(* IEC 61131-3 sources: sigmatek-logger-api/IXON_API/Class/_TCPIPClient (part 2) *)

END_FUNCTION

FUNCTION _TCPIPClient::SendTCP
	VAR_INPUT
		pConnection 	: ^_CONNECTION;
		pData 	: ^CHAR;
		udSize 	: UDINT;
		udTimeout 	: UDINT;
	END_VAR
	VAR_OUTPUT
		dRetcode 	: DINT;
	END_VAR

  dRetcode := OS_TCP_USER_SEND(pConnection^.dSocket,
                               pData,
                               udSize,
                               0, //### flags ... not used
                               udTimeout
                               );

  if (dRetcode = udSize$DINT) then
    pConnection^.udTimeStamp := ops.tAbsolute;
  else
    udSendError += 1;
    pConnection^.FSM_TCP := _STATE_SHUTDOWN;
  end_if;

END_FUNCTION

FUNCTION _TCPIPClient::SetSocketOptions
	VAR_INPUT
		dHandle 	: DINT;
	END_VAR
	VAR_OUTPUT
		Retcode 	: DINT;
	END_VAR
VAR
	OptionValue       : DINT;
  pConn             : ^_CONNECTION;
  dRet              : DINT;
  KeepAliveLasalOS  : _KeepAliveParaLasalOS;
END_VAR

  Retcode := TCP_CLT_NO_ERROR;

  if (CheckHandleValid(dHandle) = true) then

    pConn := dHandle$^_CONNECTION;

    AP_SemaWait(AP_SemaSockOpt);

    // -----------------------------------------------------------
    // - SOCKET OPTION NAGLE
    // -----------------------------------------------------------
    if (pConn^.ConnSockOpt.Nagle = true) then
      OptionValue := 1;
    else
      OptionValue := 0;
    end_if;
    dRet := OS_TCP_USER_SETSOCKOPT(pConn^.dSocket, SOL_SOCKET, SO_NAGLE, (#OptionValue)$^CHAR, sizeof(DINT));
    if (dRet < 0) then
      Retcode := dRet;
      ConnErrCallback(pConn, TCP_CLT_ERR_GROUP_OS, dRet);
    end_if;

    // -----------------------------------------------------------
    // - SOCKET OPTION KEEP ALIVE
    // -----------------------------------------------------------
    if (bdStatus.SalamanderOS = false) then
      // --------------------------------------------------------
      // - LASAL OS
      // --------------------------------------------------------
      if (pConn^.ConnSockOpt.KeepAlive = true) then
        KeepAliveLasalOS.interval := to_UINT(pConn^.KeepAlivePara.keepIDLE);
        KeepAliveLasalOS.retry    := to_UINT(pConn^.KeepAlivePara.keepINTVL);
        KeepAliveLasalOS.timeout  := to_UINT(pConn^.KeepAlivePara.keepCNT * pConn^.KeepAlivePara.keepINTVL);
      else
        KeepAliveLasalOS.interval := 0;
        KeepAliveLasalOS.retry    := 0;
        KeepAliveLasalOS.timeout  := 0;
      end_if;
      dRet := OS_TCP_USER_SETSOCKOPT(pConn^.dSocket, SOL_SOCKET, 8, (#KeepAliveLasalOS)$^CHAR, sizeof(_KeepAliveParaLasalOS));
      if (dRet < 0) then
        Retcode := dRet;
        ConnErrCallback(pConn, TCP_CLT_ERR_GROUP_OS, dRet);
      end_if;
    else
      // --------------------------------------------------------
      // - SALAMANDER OS
      // --------------------------------------------------------
      if (pConn^.ConnSockOpt.KeepAlive = true) then
        OptionValue := 1;
      else
        OptionValue := 0;
      end_if;
      dRet := OS_TCP_USER_SETSOCKOPT(pConn^.dSocket, SOL_SOCKET, 8, (#OptionValue)$^CHAR, sizeof(DINT));
      if (dRet < 0) then
        Retcode := dRet;
        ConnErrCallback(pConn, TCP_CLT_ERR_GROUP_OS, dRet);
      end_if;

//      if (pConn^.ConnSockOpt.KeepAlive = true) then
//        OptionValue := KeepAlivePara.keepCNT;
//        dRet := OS_TCP_USER_SETSOCKOPT(pConn^.dSocket, SOL_TCP, TCP_KEEPCNT, (#OptionValue)$^CHAR, sizeof(DINT));
//        if (dRet < 0) then
//          Retcode := dRet;
//          ConnErrCallback(pConn, TCP_CLT_ERR_GROUP_OS, dRet);
//        end_if;
//        OptionValue := KeepAlivePara.keepIDLE;
//        dRet := OS_TCP_USER_SETSOCKOPT(pConn^.dSocket, SOL_TCP, TCP_KEEPIDLE, (#OptionValue)$^CHAR, sizeof(DINT));
//        if (dRet < 0) then
//          Retcode := dRet;
//          ConnErrCallback(pConn, TCP_CLT_ERR_GROUP_OS, dRet);
//        end_if;
//        OptionValue := KeepAlivePara.keepINTVL;
//        dRet := OS_TCP_USER_SETSOCKOPT(pConn^.dSocket, SOL_TCP, TCP_KEEPINTVL, (#OptionValue)$^CHAR, sizeof(DINT));
//        if (dRet < 0) then
//          Retcode := dRet;
//          ConnErrCallback(pConn, TCP_CLT_ERR_GROUP_OS, dRet);
//        end_if;
//      end_if;
    end_if;

    // -----------------------------------------------------------
    // - SOCKET OPTION DELAYED ACK
    // -----------------------------------------------------------
    if (pConn^.ConnSockOpt.DelayedAck = true) then
      OptionValue := 1;
    else
      OptionValue := 0;
    end_if;
    dRet := OS_TCP_USER_SETSOCKOPT(pConn^.dSocket, SOL_SOCKET, SO_DELAYED_ACK, (#OptionValue)$^CHAR, sizeof(DINT));
    if (dRet < 0) then
      Retcode := dRet;
      ConnErrCallback(pConn, TCP_CLT_ERR_GROUP_OS, dRet);
    end_if;

    pConn^.bdSettings.SockOptChanged := false;

    AP_SemaSignal(AP_SemaSockOpt);

  else
    Retcode := TCP_CLT_INVALID_HANDLE;
  end_if;

END_FUNCTION

FUNCTION _TCPIPClient::Read_LSLOBJ_CRC32
	VAR_INPUT
		pCRC32 	: ^CHAR;
	END_VAR
	VAR_OUTPUT
		Retcode 	: DINT;
	END_VAR
VAR
	udStrLen    : UDINT;
  udCRC32     : UDINT;
  szObjName   : ARRAY [0..255] OF CHAR;
END_VAR

  Retcode := TCP_CLT_NO_ERROR;

  if (pCRC32 <> NIL) then
    pCRC32^ := 0x00;
    udStrLen := _GetObjName(this, #szObjName[0]);
    if (udStrLen > 0) then
      udCRC32 := CheckSum.CRC32(#szObjName[0], udStrLen, 0);
      SigCLib.IToA(udCRC32$DINT, pCRC32, 0x10);
    else
      Retcode := TCP_CLT_ERR_GET_LSLOBJ_NAME;
    end_if;
  else
    Retcode := TCP_CLT_ERR_INVALID_POINTER;
  end_if;

END_FUNCTION

FUNCTION _TCPIPClient::Read_AP_TaskPeriod
	VAR_OUTPUT
		Retcode 	: DINT;
	END_VAR
VAR
	dRet          : DINT;
  LSLOBJ_INFO   : LSLOBJ_INFO;
END_VAR

  Retcode := TCP_CLT_NO_ERROR;

  dRet := _TaskObjectControl.GetObjectInfo(this, OBJ_CT, #LSLOBJ_INFO);
  case dRet of
    (*=============================================================================*)
    0: // - GET OBJECT INFO OK
    (*=============================================================================*)
      if (bdStatus.SalamanderOS = true) then
        // --------------------------------------------------------
        // - SALAMANDER OS
        // --------------------------------------------------------
        if (LSLOBJ_INFO.orgperiod AND 0x80000000) then
          // -------------------------------------------------------
          // - TASK PERIOD IN [µs]
          // -------------------------------------------------------
          AP_TaskTime := LSLOBJ_INFO.orgperiod XOR 0x80000000;
        else
          // -------------------------------------------------------
          // - TASK PERIOD IN [ms]
          // -------------------------------------------------------
          AP_TaskTime := LSLOBJ_INFO.orgperiod * 1000;
        end_if;
      else
        // --------------------------------------------------------
        // - LASAL OS
        // --------------------------------------------------------
        if (LSLOBJ_INFO.orgperiod AND 0x80000000) then
          // -------------------------------------------------------
          // - TASK PERIOD IN [µs]
          // -------------------------------------------------------
          AP_TaskTime := (LSLOBJ_INFO.orgperiod XOR 0x80000000) / 1000;
          if (AP_TaskTime = 0) then
            AP_TaskTime := 1;
          end_if;
        else
          // -------------------------------------------------------
          // - TASK PERIOD IN [ms]
          // -------------------------------------------------------
          AP_TaskTime := LSLOBJ_INFO.orgperiod;
        end_if;
      end_if;

    (*=============================================================================*)
    -1: // - ERROR READ OBJECT INFO (NO APPLICATION)
    (*=============================================================================*)
      Retcode     := TCP_CLT_ERR_TASK_TIME_NO_APP;
      AP_TaskTime := 0xFFFFFFFF;

    (*=============================================================================*)
    -3: // - ERROR READ OBJECT INFO (NO APPLICATION)
    (*=============================================================================*)
      Retcode     := TCP_CLT_ERR_TASK_TIME_WRONG_TASK_TYPE;
      AP_TaskTime := 0xFFFFFFFF;

    (*=============================================================================*)
    -5: // - OBJECT NOT FOUND (TASK DEACTIVATED)
    (*=============================================================================*)
      Retcode     := TCP_CLT_ERR_TASK_TIME_OBJ_NOT_FOUND;
      AP_TaskTime := 0xFFFFFFFF;

  end_case;

END_FUNCTION

FUNCTION _TCPIPClient::GetMultiTaskErrorCode
	VAR_INPUT
		pErrTxt 	: ^CHAR;
	END_VAR
VAR
	ErrMT     : DINT;
END_VAR

  ErrMT := _MultiTask.GETLASTERROR();
  case ErrMT of

    (*===============================================================================================*)
    MTERROR_NONE: // - NO ERROR
    (*===============================================================================================*)
      SigCLib.StrCpy(pErrTxt, "MTERROR_NONE");

    (*===============================================================================================*)
    MTERROR_NOMEM: // - NO MORE MEMORY TO RUN THIS FUNCTION, E.G. INTERNAL ALLOC FAILED
    (*===============================================================================================*)
      SigCLib.StrCpy(pErrTxt, "MTERROR_NOMEM");

    (*===============================================================================================*)
    MTERROR_NOFCT: // - CREATE TASK NEEDS A VALID TASK FUNCTION
    (*===============================================================================================*)
      SigCLib.StrCpy(pErrTxt, "MTERROR_NOFCT");

    (*===============================================================================================*)
    MTERROR_FCTNOTINMEM: // - CREATE TASK NEEDS A TASK FUNCTION PLACED IN LASAL CODE MEMORY
    (*===============================================================================================*)
      SigCLib.StrCpy(pErrTxt, "MTERROR_FCTNOTINMEM");

    (*===============================================================================================*)
    MTERROR_WRONGPRIOR: // - CREATE TASK ONLY SUPPORTS PRIORS FROM 1 .. 14
    (*===============================================================================================*)
      SigCLib.StrCpy(pErrTxt, "MTERROR_WRONGPRIOR");

    (*===============================================================================================*)
    MTERROR_STACK: // - CREATE TASK ONLY SUPPORT SATCK SIZE LOWER THAN 0x4000
    (*===============================================================================================*)
      SigCLib.StrCpy(pErrTxt, "MTERROR_STACK");

    (*===============================================================================================*)
    MTERROR_NAME: // - CREATE TASK, MAILBOX OR SEMAPHORE NEEDS A VALID NAME
    (*===============================================================================================*)
      SigCLib.StrCpy(pErrTxt, "MTERROR_NAME");

    (*===============================================================================================*)
    MTERROR_NAMEUSED: // - CREATE TASK, MAILBOX OR SEMAPHORE NAME ALREADY IN USE
    (*===============================================================================================*)
      SigCLib.StrCpy(pErrTxt, "MTERROR_NAMEUSED");

    (*===============================================================================================*)
    MTERROR_HANDLE: // - HANDLE NOT FOUND IN OS-LIST => NOT VALID
    (*===============================================================================================*)
      SigCLib.StrCpy(pErrTxt, "MTERROR_HANDLE");

    (*===============================================================================================*)
    MTERROR_NOTALLOWED: // - MT-FUNCTION NOT ALLOWED IN THIS TASK CONTEXT
    (*===============================================================================================*)
      SigCLib.StrCpy(pErrTxt, "MTERROR_NOTALLOWED");

    (*===============================================================================================*)
    MTERROR_MESSAGESIZE: // - MAILBOX NEED A VALID MESSAGE SIZE
    (*===============================================================================================*)
      SigCLib.StrCpy(pErrTxt, "MTERROR_MESSAGESIZE");

    (*===============================================================================================*)
    MTERROR_DATA: // - POINTER TO DATA IS NOT VALID
    (*===============================================================================================*)
      SigCLib.StrCpy(pErrTxt, "MTERROR_DATA");

    (*===============================================================================================*)
    MTERROR_PTR: // - INVALID POINTER, PARAMETER OR INTERNAL
    (*===============================================================================================*)
      SigCLib.StrCpy(pErrTxt, "MTERROR_PTR");

    (*===============================================================================================*)
    MTERROR_TASKID: // - INVALID TASK ID, ID NOT FOUND
    (*===============================================================================================*)
      SigCLib.StrCpy(pErrTxt, "MTERROR_TASKID");

    (*===============================================================================================*)
    MTERROR_NOTASK: // - TASK DOES NOT EXIST
    (*===============================================================================================*)
      SigCLib.StrCpy(pErrTxt, "MTERROR_NOTASK");

    (*===============================================================================================*)
    MTERROR_NOIFFNC: // - INTERFACE FUNCTION IS NOT AVAILABLE
    (*===============================================================================================*)
      SigCLib.StrCpy(pErrTxt, "MTERROR_NOIFFNC");

    (*===============================================================================================*)
    else // - UNKNOWN ERROR CODE
    (*===============================================================================================*)
      SigCLib.StrCpy(pErrTxt, "MTERROR_UNKNOWN");

  end_case;

END_FUNCTION

FUNCTION _TCPIPClient::AP_TaskCreate
	VAR_INPUT
		pTaskName 	: ^CHAR;
		pCallback 	: ^void;
	END_VAR
	VAR_OUTPUT
		Retcode 	: DINT;
	END_VAR

  Retcode := TCP_CLT_NO_ERROR;

  AP_TaskHandle := _MultiTask.CREATETHREAD(pCallback, AP_TaskPriority, 0x4000, MT_TASK_SAVETHIS, this, pTaskName);
  if (AP_TaskHandle = NIL) then
    Retcode := TCP_CLT_ERR_TASK_CREATE;
  end_if;

END_FUNCTION

FUNCTION __CDECL _TCPIPClient::AP_TaskCallback
	VAR_INPUT
		Param0 	: ^void;
	END_VAR

  while 1 do
    CyclicCall();
    AP_TaskDelay(AP_TaskTime);
  end_while;

END_FUNCTION

FUNCTION _TCPIPClient::AP_TaskDelay
	VAR_INPUT
		udTaskDelay 	: UDINT;
	END_VAR

  if (bdStatus.SalamanderOS = true) then
    OSSD_DELAY(pCIL_DEBUG, udTaskDelay);
  else
    _MultiTask.TASKDELAY(udTaskDelay);
  end_if;

END_FUNCTION

FUNCTION _TCPIPClient::AP_SemaCreate
	VAR_INPUT
		pSemaName 	: ^CHAR;
		Index 	: DINT;
	END_VAR
	VAR_OUTPUT
		Retcode 	: DINT;
	END_VAR

  Retcode := TCP_CLT_NO_ERROR;

  if (pSemaName <> NIL) then
    case Index of
      (*=================================================================================*)
      0:
      (*=================================================================================*)
        AP_SemaHandle1 := _MultiTask.CREATESEMAPHORE(MTSEMATYPE_MUTEX, 1, 0, pSemaName);
        if (AP_SemaHandle1 = NIL) then
          Retcode := TCP_CLT_ERR_SEMA_CREATE;
        end_if;

      (*=================================================================================*)
      1:
      (*=================================================================================*)
        AP_SemaSockOpt := _MultiTask.CREATESEMAPHORE(MTSEMATYPE_MUTEX, 1, 0, pSemaName);
        if (AP_SemaSockOpt = NIL) then
          Retcode := TCP_CLT_ERR_SEMA_CREATE;
        end_if;

      (*=================================================================================*)
      else
      (*=================================================================================*)
        Retcode := TCP_CLT_ERR_SEMA_INVALID_IDX;

    end_case;
  else
    Retcode := TCP_CLT_ERR_SEMA_INVALID_NAME;
  end_if;

END_FUNCTION

FUNCTION _TCPIPClient::AP_SemaWait
	VAR_INPUT
		SemaHandle 	: MT_SEMAHANDLE;
	END_VAR

  if (SemaHandle <> NIL) then
    _MultiTask.WAIT(SemaHandle);
  end_if;

END_FUNCTION

FUNCTION _TCPIPClient::AP_SemaSignal
	VAR_INPUT
		SemaHandle 	: MT_SEMAHANDLE;
	END_VAR

  if (SemaHandle <> NIL) then
    _MultiTask.SIGNAL(SemaHandle);
  end_if;

END_FUNCTION

FUNCTION _TCPIPClient::DelConnIntern
	VAR_INPUT
		pDelConn 	: ^_CONNECTION;
	END_VAR
VAR
	pSearchConn : ^_CONNECTION;
END_VAR

  if (pDelConn <> NIL) then

    AP_SemaWait(AP_SemaHandle1);

    if (pDelConn^.pNextConn = pDelConn) then
      // - ONE ACTIVE CONNECTION
    else
      pSearchConn := pDelConn;
      while pSearchConn^.pNextConn <> pDelConn do
        pSearchConn := pSearchConn^.pNextConn;
      end_while;
      pSearchConn^.pNextConn := pDelConn^.pNextConn;
      pActConn := pDelConn^.pNextConn;
      bdStatus.InhibNextConn := true;
    end_if;

    ConnInfoCallback(pDelConn, TCP_CLT_INFO_DELETED, 0);
    INITConnection(pDelConn);
    AP_SemaSignal(AP_SemaHandle1);

    ActConn -= 1;

  end_if;

END_FUNCTION

FUNCTION _TCPIPClient::AddConnIntern
	VAR_INPUT
		pIPAddress 	: ^CHAR;
		pCACertPEMFilename 	: ^CHAR;
		pClientCertChainPEMFilename 	: ^CHAR;
		pClientCertKeyPEMFilename 	: ^CHAR;
		pKeyDecryptPwd 	: ^CHAR;
		pCallbackThis 	: ^_TCPIPClientInterface;
		udTimeout 	: UDINT;
		ConnSSL 	: BOOL;
	END_VAR
	VAR_OUTPUT
		dHandle 	: DINT;
	END_VAR
VAR
  pFirstConn                    : ^_CONNECTION;
  pNewConn                      : ^_CONNECTION;
  pSearchConn                   : ^_CONNECTION;
  i                             : USINT;
END_VAR

  dHandle := 0;

  if (pIPAddress = NIL) | (pConnectionBuffer = NIL) | (Control = _STATE_ERROR_CREATING_MUTEX) | (Control = _STATE_ERROR_ALLOCATING_MEMORY) then
    return;
  end_if;

  if (ActConn < MaxConn) then

    AP_SemaWait(AP_SemaHandle1);

    for i := 0 to (MaxConn-1) do
      pFirstConn := pConnectionBuffer + (i * sizeof(_CONNECTION));
      if (pFirstConn^.bInUse = true) then
        exit;
      else
        pFirstConn := NIL;
      end_if;
    end_for;

    for i := 0 to (MaxConn-1) do
      pNewConn := pConnectionBuffer + (i * sizeof(_CONNECTION));
      if (pNewConn^.bInUse = false) then
        exit;
      end_if;
    end_for;

    pNewConn^.bInUse          := true;
    pNewConn^.udTimeout       := udTimeout;
    pNewConn^.pCallbackThis   := pCallbackThis;
    pNewConn^.FSM_TCP         := _STATE_IDLE;
    pNewConn^.ConnSockOpt     := MainSockOpt;
    pNewConn^.KeepAlivePara   := KeepAlivePara;
    pNewConn^.CloseSocketType := CloseSocketType;
    SigCLib.StrCpy(#pNewConn^.szIPAddress[0], pIPAddress);
    pNewConn^.bdSettings.SockOptChanged := true;

    if (ConnSSL = true) then
      pNewConn^.bdSettings.ConnSSL := true;
      if (pCACertPEMFilename <> NIL) then
        SigCLib.StrCpy(#pNewConn^.szCACertPEMFileName[0], pCACertPEMFilename);
      end_if;
      if (pClientCertChainPEMFilename <> NIL) then
        SigCLib.StrCpy(#pNewConn^.szClientCertChainPEMFilename[0], pClientCertChainPEMFilename);
      end_if;
      if (pClientCertKeyPEMFilename <> NIL) then
        SigCLib.StrCpy(#pNewConn^.szClientCertKeyPEMFilename[0], pClientCertKeyPEMFilename);
      end_if;
      if (pKeyDecryptPwd <> NIL) then
        SigCLib.StrCpy(#pNewConn^.szKeyDecryptPwd[0], pKeyDecryptPwd);
      end_if;
    end_if;

    if (pFirstConn = NIL) then
      pNewConn^.pNextConn := pNewConn;
    else
      pSearchConn := pFirstConn;
      while (pSearchConn^.pNextConn <> pFirstConn) do
        pSearchConn := pSearchConn^.pNextConn;
      end_while;
      pNewConn^.pNextConn    := pFirstConn;
      pSearchConn^.pNextConn := pNewConn;
    end_if;

    dHandle := pNewConn$DINT;
    ActConn += 1;

    AP_SemaSignal(AP_SemaHandle1);

  else
    LastError := TCP_CLT_ERR_MAX_CONN;
  end_if;

END_FUNCTION

FUNCTION _TCPIPClient::CheckParaConnSSL
	VAR_INPUT
		pCACertPEMFilename 	: ^CHAR;
		pClientCertChainPEMFilename 	: ^CHAR;
		pClientCertKeyPEMFilename 	: ^CHAR;
		pKeyDecryptPwd 	: ^CHAR;
	END_VAR
	VAR_OUTPUT
		Retcode 	: DINT;
	END_VAR

  Retcode := TCP_CLT_NO_ERROR;

  if (pClientCertChainPEMFilename <> NIL) then
    if (pClientCertKeyPEMFilename = NIL) then
      Retcode := TCP_CLT_ERR_INVALID_PARA_SSL;
    end_if;
  end_if;

  if (pClientCertKeyPEMFilename <> NIL) then
    if (pClientCertChainPEMFilename = NIL) then
      Retcode := TCP_CLT_ERR_INVALID_PARA_SSL;
    end_if;
  end_if;

  if (pKeyDecryptPwd <> NIL) then
    if (pClientCertChainPEMFilename = NIL) then
      Retcode := TCP_CLT_ERR_INVALID_PARA_SSL;
    end_if;
    if (pClientCertKeyPEMFilename = NIL) then
      Retcode := TCP_CLT_ERR_INVALID_PARA_SSL;
    end_if;
  end_if;

END_FUNCTION

FUNCTION _TCPIPClient::FindFirstConn
	VAR_OUTPUT
		pFirstConn 	: ^_CONNECTION;
	END_VAR
VAR
	i           : USINT;
  pSearchConn : ^_CONNECTION;
END_VAR

  pFirstConn := NIL;

  for i := 0 to (MaxConn-1) do
    pSearchConn := pConnectionBuffer + (i * sizeof(_CONNECTION));
    if (pSearchConn^.bInUse = true) then
      pFirstConn := pSearchConn;
    end_if;
  end_for;

END_FUNCTION

FUNCTION _TCPIPClient::CheckParaConnTCP
	VAR_INPUT
		pIPAddress 	: ^CHAR;
		pCallbackThis 	: ^void;
	END_VAR
	VAR_OUTPUT
		Retcode 	: DINT;
	END_VAR
VAR
	udStrLen        : UDINT;
END_VAR

  Retcode := TCP_CLT_NO_ERROR;

  if (pIPAddress = NIL) then
    Retcode := TCP_CLT_ERR_INVALID_PARA_TCP;
  else
    udStrLen := SigCLib.StrLen(pIPAddress);
    if (udStrLen = 0) then
      Retcode := TCP_CLT_ERR_INVALID_PARA_TCP;
    end_if;
  end_if;

  if (pCallbackThis = NIL) then
    Retcode := TCP_CLT_ERR_INVALID_PARA_TCP;
  end_if;

END_FUNCTION

FUNCTION _TCPIPClient::ConnErrCallback
	VAR_INPUT
		pConn 	: ^_CONNECTION;
		ErrGroup 	: DINT;
		ErrCode 	: DINT;
	END_VAR
	VAR_OUTPUT
		Retcode 	: DINT;
	END_VAR

  Retcode := TCP_CLT_NO_ERROR;

  if (pConn <> NIL) then
    if (pConn^.pCallbackThis <> NIL) then
      pConn^.pCallbackThis$^_TCPIPClientInterface^.ErrCallback(pConn^.FSM_TCP, ErrGroup, ErrCode);
    end_if;
  else
    Retcode := TCP_CLT_INVALID_HANDLE;
  end_if;

END_FUNCTION
FUNCTION _TCPIPClient::ConnInfoCallback
	VAR_INPUT
		pConn 	: ^_CONNECTION;
		InfoPara1 	: DINT;
		InfoPara2 	: DINT;
	END_VAR
	VAR_OUTPUT
		Retcode 	: DINT;
	END_VAR

  Retcode := TCP_CLT_NO_ERROR;

  if (pConn <> NIL) then
    if (pConn^.pCallbackThis <> NIL) then
      pConn^.pCallbackThis$^_TCPIPClientInterface^.InfoCallback(pConn^.FSM_TCP, InfoPara1, InfoPara2);
    end_if;
  else
    Retcode := TCP_CLT_INVALID_HANDLE;
  end_if;

END_FUNCTION
FUNCTION _TCPIPClient::AP_NReadAvailable
	VAR_INPUT
		pConn 	: ^_CONNECTION;
	END_VAR
	VAR_OUTPUT
		Retcode 	: DINT;
	END_VAR

  if (pConn <> NIL) then
    if (pConn^.bdSettings.ConnSSL = false) then
      Retcode := OS_TCP_USER_NREAD_AVAILABLE(pConn^.dSocket);
    else
      Retcode := SizeOfTXBuffer$DINT;
    end_if;
  else
    Retcode := TCP_CLT_INVALID_HANDLE;
  end_if;

END_FUNCTION

FUNCTION _TCPIPClient::INITConnection
	VAR_INPUT
		pConnection 	: ^_CONNECTION;
	END_VAR

  pConnection^.bInUse     := false;
  pConnection^.bConnected := false;
  pConnection^.dSocket    := 0;
  pConnection^.FSM_TCP    := _STATE_IDLE;

  pConnection^.pCallbackThis := NIL;

  pConnection^.udTimeout   := 0;
  pConnection^.udTimeStamp := 0;

  pConnection^.RingbufferForSending.udUsed := 0;
  pConnection^.RingbufferForSending.pRead  := pConnection^.RingbufferForSending.pMem;
  pConnection^.RingbufferForSending.pWrite := pConnection^.RingbufferForSending.pMem;
  pConnection^.BufferHeader.DataSize       := 0;
  pConnection^.pSendReceiveBufferHelp      := pConnection^.pSendReceiveBuffer;

  pConnection^.ConnSockOpt := MainSockOpt;
  pConnection^.pNextConn   := NIL;

  pConnection^.bdSettings.DelConn        := false;
  pConnection^.bdSettings.ConnSSL        := false;
  pConnection^.bdSettings.SockOptChanged := false;

  SigCLib.MemSet(#pConnection^.szIPAddress[0], 0x00, 0x10);
  SigCLib.MemSet(#pConnection^.szCACertPEMFilename, 0x00, sizeof(_CONNECTION.szCACertPEMFilename));
  SigCLib.MemSet(#pConnection^.szClientCertChainPEMFilename, 0x00, sizeof(_CONNECTION.szClientCertChainPEMFilename));
  SigCLib.MemSet(#pConnection^.szClientCertKeyPEMFilename, 0x00, sizeof(_CONNECTION.szClientCertKeyPEMFilename));
  SigCLib.MemSet(#pConnection^.szKeyDecryptPwd, 0x00, sizeof(_CONNECTION.szKeyDecryptPwd));

  pConnection^.KeepAlivePara   := KeepAlivePara;
  pConnection^.CloseSocketType := CloseSocketType;

END_FUNCTION

FUNCTION _TCPIPClient::SendSSL
	VAR_INPUT
		pConnection 	: ^_CONNECTION;
		pData 	: ^CHAR;
		udSize 	: UDINT;
		udTimeout 	: UDINT;
	END_VAR
	VAR_OUTPUT
		dRetcode 	: DINT;
	END_VAR

  dRetcode := OS_SSL_USER_WRITE(pConnection^.dSocket,
                                pData,
                                to_dint(udSize),
                                udTimeout);

  if (dRetcode = udSize$DINT) then
    pConnection^.udTimeStamp := ops.tAbsolute;
  else
    udSendError += 1;
    pConnection^.FSM_TCP := _STATE_SHUTDOWN;
  end_if;

END_FUNCTION
